// TIA Portal V20 export
TextList "TextList_ScreenNames"  ListRange=Decimal
  TextListEntry   EntryType=SingleValue, From=1, To=1, Text="Root screen"
